FUNCTION_BLOCK FB_Event_echo // for HMI event pudate purpose
VAR_INPUT
END_VAR
VAR_OUTPUT
	echo: INT;
END_VAR
VAR
	ton_time: TON;
	Puls: INT;
	
	memo: BOOL;

END_VAR

ton_time(PT:=T#2S,IN:=memo AND NOT ton_time.Q);
IF ton_time.Q THEN;
	echo:=echo+1;
	
	IF Puls>=5 THEN;
		memo:=FALSE;
	ELSE;
		Puls:=Puls+1;
	END_IF
END_IF

IF ton_time.Q THEN;
	ton_time.IN:=FALSE;
END_IF

METHOD event : BOOL
VAR_INPUT
END_VAR
memo:=TRUE;
echo:=0;
Puls:=0;
END_METHOD

END_FUNCTION_BLOCK

(* stored: Version 1.1.0.1, ProductVersion 3.1.4024.15
   POU FB_Event_echo: Id {8e4667bf-577c-479e-878c-e91bfc8e7d87}, SpecialFunc None
   Method event: Id {1489a449-054b-4248-87c6-4ec2e3069a24} *)
